// TIA Portal V20 export
Screen "Sew_TurnTable"  1276x673
  ScreenItem "Rectangle_5" at 197,72 size 248x590  Type=HmiRectangle
  ScreenItem "Rectangle_3" at 451,72 size 248x585  Type=HmiRectangle
  ScreenItem "符号 IO 域_7" at 390,6 size 500x41  Type=HmiSymbolicIOField
  ScreenItem "permanentareaborderrectangle" at 0,0 size 0x0  Type=HmiRectangle
  ScreenItem "Line_Header_X0_Y64" at 0,65 size 1280x0  Type=HmiLine
  ScreenItem "Button_Back" at 2,2 size 90x60  Type=HmiButton
  ScreenItem "Text_DigitalOutputs_30" at 519,134 size 124x16  Type=HmiTextBox
  ScreenItem "Text_DigitalOutputs_31" at 519,158 size 124x16  Type=HmiTextBox
  ScreenItem "Text_DigitalOutputs_32" at 519,182 size 124x16  Type=HmiTextBox
  ScreenItem "Text_DigitalOutputs_34" at 519,207 size 124x16  Type=HmiTextBox
  ScreenItem "Text_DigitalOutputs_35" at 519,231 size 124x16  Type=HmiTextBox
  ScreenItem "LED_1_Left_33" at 0,0 size 100x30  Type=HmiCircle
  ScreenItem "LED_1_Left_23" at 0,0 size 100x30  Type=HmiCircle
  ScreenItem "LED_1_Left_24" at 0,0 size 100x30  Type=HmiCircle
  ScreenItem "LED_1_Left_25" at 0,0 size 100x30  Type=HmiCircle
  ScreenItem "LED_1_Left_26" at 0,0 size 100x30  Type=HmiCircle
  ScreenItem "按钮_5" at 202,562 size 115x72  Type=HmiButton
  ScreenItem "按钮_8" at 320,562 size 115x72  Type=HmiButton
  ScreenItem "按钮_9" at 202,395 size 115x72  Type=HmiButton
  ScreenItem "按钮_10" at 323,395 size 115x72  Type=HmiButton
  ScreenItem "按钮_3" at 459,561 size 115x72  Type=HmiButton
  ScreenItem "按钮_2" at 459,486 size 115x72  Type=HmiButton
  ScreenItem "按钮_1" at 459,412 size 115x72  Type=HmiButton
  ScreenItem "按钮_7" at 459,338 size 115x72  Type=HmiButton
  ScreenItem "IO 域_9" at 576,338 size 115x72  Type=HmiIOField
  ScreenItem "文本_1" at 470,314 size 94x24  Type=HmiText
  ScreenItem "文本_2" at 587,314 size 94x24  Type=HmiText
  ScreenItem "IO 域_10" at 576,412 size 115x72  Type=HmiIOField
  ScreenItem "IO 域_11" at 576,486 size 115x72  Type=HmiIOField
  ScreenItem "IO 域_12" at 576,561 size 115x72  Type=HmiIOField
  ScreenItem "文本_3" at 207,130 size 94x24  Type=HmiText
  ScreenItem "IO 域_13" at 305,122 size 116x39  Type=HmiIOField
  ScreenItem "文本_4" at 207,170 size 94x24  Type=HmiText
  ScreenItem "IO 域_14" at 305,162 size 116x39  Type=HmiIOField
  ScreenItem "按钮_11" at 202,203 size 115x72  Type=HmiButton
  ScreenItem "按钮_12" at 202,319 size 115x72  Type=HmiButton
  ScreenItem "按钮_6" at 199,73 size 498x40  Type=HmiButton
  ScreenItem "Rectangle_4" at 9,64 size 180x273  Type=HmiRectangle
  ScreenItem "Graphic view_1" at 14,75 size 61x38  Type=HmiGraphicView
  ScreenItem "Graphic view_2" at 124,75 size 61x38  Type=HmiGraphicView
  ScreenItem "Text_DigitalOutputs_33" at 16,120 size 91x16  Type=HmiTextBox
  ScreenItem "LED_1_Left_1" at 0,0 size 100x30  Type=HmiCircle
  ScreenItem "Text_DigitalOutputs_1" at 29,209 size 100x16  Type=HmiTextBox
  ScreenItem "IO 域_1" at 110,117 size 54x21  Type=HmiIOField
  ScreenItem "IO 域_2" at 110,139 size 54x21  Type=HmiIOField
  ScreenItem "IO 域_3" at 110,161 size 54x21  Type=HmiIOField
  ScreenItem "IO 域_4" at 110,183 size 54x21  Type=HmiIOField
  ScreenItem "Text_DigitalOutputs_2" at 16,142 size 91x16  Type=HmiTextBox
  ScreenItem "Text_DigitalOutputs_3" at 16,164 size 91x16  Type=HmiTextBox
  ScreenItem "Text_DigitalOutputs_4" at 16,186 size 91x16  Type=HmiTextBox
  ScreenItem "Text_DigitalOutputs_5" at 29,225 size 100x16  Type=HmiTextBox
  ScreenItem "Text_DigitalOutputs_6" at 29,258 size 100x16  Type=HmiTextBox
  ScreenItem "Text_DigitalOutputs_7" at 29,274 size 100x16  Type=HmiTextBox
  ScreenItem "Text_DigitalOutputs_8" at 29,291 size 100x16  Type=HmiTextBox
  ScreenItem "Text_DigitalOutputs_9" at 29,307 size 100x16  Type=HmiTextBox
  ScreenItem "Text_DigitalOutputs_10" at 29,324 size 100x16  Type=HmiTextBox
  ScreenItem "Text_DigitalOutputs_11" at 29,241 size 100x16  Type=HmiTextBox
  ScreenItem "LED_1_Left_2" at 0,0 size 100x30  Type=HmiCircle
  ScreenItem "LED_1_Left_3" at 0,0 size 100x30  Type=HmiCircle
  ScreenItem "LED_1_Left_4" at 0,0 size 100x30  Type=HmiCircle
  ScreenItem "LED_1_Left_5" at 0,0 size 100x30  Type=HmiCircle
  ScreenItem "LED_1_Left_6" at 0,0 size 100x30  Type=HmiCircle
  ScreenItem "LED_1_Left_7" at 0,0 size 100x30  Type=HmiCircle
  ScreenItem "LED_1_Left_8" at 0,0 size 100x30  Type=HmiCircle
  ScreenItem "线_1" at 76,95 size 45x0  Type=HmiLine
  ScreenItem "Rectangle_1" at 9,337 size 180x335  Type=HmiRectangle
  ScreenItem "Text_DigitalOutputs_12" at 33,442 size 108x16  Type=HmiTextBox
  ScreenItem "Text_DigitalOutputs_13" at 33,458 size 108x16  Type=HmiTextBox
  ScreenItem "Text_DigitalOutputs_14" at 33,474 size 108x16  Type=HmiTextBox
  ScreenItem "Text_DigitalOutputs_20" at 33,491 size 108x16  Type=HmiTextBox
  ScreenItem "Text_DigitalOutputs_21" at 33,507 size 108x16  Type=HmiTextBox
  ScreenItem "Text_DigitalOutputs_22" at 33,524 size 108x16  Type=HmiTextBox
  ScreenItem "Text_DigitalOutputs_23" at 33,540 size 108x16  Type=HmiTextBox
  ScreenItem "Text_DigitalOutputs_24" at 33,557 size 108x16  Type=HmiTextBox
  ScreenItem "Text_DigitalOutputs_25" at 33,573 size 108x16  Type=HmiTextBox
  ScreenItem "Text_DigitalOutputs_26" at 33,590 size 108x16  Type=HmiTextBox
  ScreenItem "Text_DigitalOutputs_27" at 33,606 size 108x16  Type=HmiTextBox
  ScreenItem "Text_DigitalOutputs_28" at 33,623 size 108x16  Type=HmiTextBox
  ScreenItem "Text_DigitalOutputs_29" at 33,639 size 108x16  Type=HmiTextBox
  ScreenItem "Text_DigitalOutputs_44" at 13,385 size 73x16  Type=HmiTextBox
  ScreenItem "IO 域_5" at 110,382 size 54x21  Type=HmiIOField
  ScreenItem "IO 域_6" at 110,404 size 54x21  Type=HmiIOField
  ScreenItem "IO 域_7" at 110,426 size 54x21  Type=HmiIOField
  ScreenItem "Text_DigitalOutputs_45" at 13,407 size 73x16  Type=HmiTextBox
  ScreenItem "Text_DigitalOutputs_46" at 13,429 size 73x16  Type=HmiTextBox
  ScreenItem "Text_DigitalOutputs_47" at 33,656 size 108x16  Type=HmiTextBox
  ScreenItem "LED_1_Left_9" at 0,0 size 100x30  Type=HmiCircle
  ScreenItem "LED_1_Left_10" at 0,0 size 100x30  Type=HmiCircle
  ScreenItem "LED_1_Left_11" at 0,0 size 100x30  Type=HmiCircle
  ScreenItem "LED_1_Left_12" at 0,0 size 100x30  Type=HmiCircle
  ScreenItem "LED_1_Left_13" at 0,0 size 100x30  Type=HmiCircle
  ScreenItem "LED_1_Left_14" at 0,0 size 100x30  Type=HmiCircle
  ScreenItem "LED_1_Left_15" at 0,0 size 100x30  Type=HmiCircle
  ScreenItem "LED_1_Left_16" at 0,0 size 100x30  Type=HmiCircle
  ScreenItem "LED_1_Left_17" at 0,0 size 100x30  Type=HmiCircle
  ScreenItem "LED_1_Left_18" at 0,0 size 100x30  Type=HmiCircle
  ScreenItem "LED_1_Left_19" at 0,0 size 100x30  Type=HmiCircle
  ScreenItem "LED_1_Left_20" at 0,0 size 100x30  Type=HmiCircle
  ScreenItem "LED_1_Left_21" at 0,0 size 100x30  Type=HmiCircle
  ScreenItem "LED_1_Left_22" at 0,0 size 100x30  Type=HmiCircle
  ScreenItem "线_2" at 80,358 size 44x1  Type=HmiLine
  ScreenItem "Graphic view_3" at 125,340 size 61x38  Type=HmiGraphicView
  ScreenItem "Graphic view_4" at 14,340 size 61x38  Type=HmiGraphicView
  ScreenItem "LED_1_Left_30" at 0,0 size 100x30  Type=HmiCircle
  ScreenItem "LED_1_Left_29" at 0,0 size 100x30  Type=HmiCircle
  ScreenItem "LED_1_Left_28" at 0,0 size 100x30  Type=HmiCircle
  ScreenItem "LED_1_Left_27" at 0,0 size 100x30  Type=HmiCircle
  ScreenItem "线_3" at 199,310 size 242x0  Type=HmiLine
  ScreenItem "线_4" at 199,491 size 241x0  Type=HmiLine
  ScreenItem "线_7" at 453,285 size 242x0  Type=HmiLine
  ScreenItem "Zone01" at 706,68 size 569x585  Type=HmiGraphicView
  ScreenItem "LED_1_Left_34" at 0,0 size 100x30  Type=HmiCircle
  ScreenItem "文本域_7" at 1029,150 size 119x33  Type=HmiTextBox
  ScreenItem "Line_1V1_4" at 1021,210 size 9x149  Type=HmiLine
  ScreenItem "文本域_1" at 731,576 size 119x33  Type=HmiTextBox
  ScreenItem "文本域_2" at 713,202 size 119x33  Type=HmiTextBox
  ScreenItem "文本域_3" at 1130,474 size 119x33  Type=HmiTextBox
  ScreenItem "Line_1V1_1" at 771,286 size 139x71  Type=HmiLine
  ScreenItem "Line_1V1_3" at 1074,483 size 55x25  Type=HmiLine
  ScreenItem "Line_1V1_5" at 780,500 size 72x87  Type=HmiLine
